(* IEC 61131-3 sources: llm-plc-st-eval/data/definitivo/qwen2.5-coder_14b/A4/few_shot, 3 files *)

(* ---- ejec_1.st ---- *)
FUNCTION_BLOCK FB_Rampa
VAR_INPUT
    SPvel : REAL; (* Consigna de velocidad *)
    paroRapido : BOOL; (* Paro rápido activo *)
    ciclo : TIME; (* Ciclo de ejecución *)
END_VAR
VAR_OUTPUT
    CVvel : REAL; (* Consigna de velocidad variable *)
END_VAR
VAR
    error : REAL; (* Error entre SPvel y CVvel *)
    dt : TIME; (* Tiempo transcurrido desde la última iteración *)
    dt_sec : REAL; (* Tiempo transcurrido en segundos *)
    rampaSubida : REAL := 10.0; (* Pendiente de subida en puntos porcentuales por segundo *)
    rampaBajada : REAL := 20.0; (* Pendiente de bajada en puntos porcentuales por segundo *)
    rampaParoRapido : REAL := 40.0; (* Pendiente de paro rápido en puntos porcentuales por segundo *)
    lastTime : TIME; (* Tiempo de la última iteración *)
END_VAR

(* Calcula el tiempo transcurrido desde la última iteración *)
dt := ciclo;
dt_sec := dt / T#1S;

(* Actualiza CVvel según las condiciones *)
IF paroRapido THEN
    (* Paro rápido activo *)
    CVvel := CVvel - rampaParoRapido * dt_sec;
    IF CVvel < 0.0 THEN
        CVvel := 0.0;
    END_IF;
ELSE
    (* Paro rápido inactivo *)
    error := SPvel - CVvel;
    IF error > 0 THEN
        (* Subida *)
        CVvel := CVvel + rampaSubida * dt_sec;
        IF CVvel > SPvel THEN
            CVvel := SPvel;
        END_IF;
    ELSE
        (* Bajada *)
        CVvel := CVvel - rampaBajada * dt_sec;
        IF CVvel < SPvel THEN
            CVvel := SPvel;
        END_IF;
    END_IF;
END_IF;

(* Actualiza el tiempo de la última iteración *)
lastTime := lastTime + ciclo;
END_FUNCTION_BLOCK

(* ---- ejec_2.st ---- *)
FUNCTION_BLOCK FB_Rampa
VAR_INPUT
    SPvel : REAL; (* Consigna de velocidad *)
    paroRapido : BOOL; (* Paro rápido activo *)
    ciclo : TIME; (* Ciclo de ejecución *)
END_VAR
VAR_OUTPUT
    CVvel : REAL; (* Condicional de velocidad *)
END_VAR
VAR
    error : REAL; (* Error entre SPvel y CVvel *)
    dt : TIME; (* Tiempo transcurrido desde la última ejecución *)
    dtSec : REAL; (* Tiempo transcurrido en segundos *)
    rampaSubida : REAL; (* Pendiente de subida *)
    rampaBajada : REAL; (* Pendiente de bajada *)
    rampaParoRapido : REAL; (* Pendiente de paro rápido *)
END_VAR

(* Inicialización de las rampas *)
rampaSubida := 10.0;
rampaBajada := 20.0;
rampaParoRapido := 40.0;

(* Cálculo del tiempo transcurrido en segundos *)
dt := ciclo;
dtSec := dt / T#1S;

(* Lógica de paro rápido *)
IF paroRapido THEN
    CVvel := MAX(0.0, CVvel - rampaParoRapido * dtSec);
ELSE
    (* Cálculo del error *)
    error := SPvel - CVvel;

    (* Ajuste de CVvel con rampa *)
    IF error > 0 THEN
        CVvel := MIN(CVvel + rampaSubida * dtSec, SPvel);
    ELSE
        CVvel := MAX(CVvel - rampaBajada * dtSec, SPvel);
    END_IF;
END_IF;

(* Evitar sobrepaso *)
IF CVvel > SPvel THEN
    CVvel := SPvel;
ELSIF CVvel < 0.0 THEN
    CVvel := 0.0;
END_IF;

END_FUNCTION_BLOCK

(* ---- ejec_3.st ---- *)
FUNCTION_BLOCK FB_Rampa
VAR_INPUT
    SPvel : REAL; (* Consigna de velocidad *)
    paroRapido : BOOL; (* Paro rápido activo *)
    ciclo : TIME; (* Ciclo de ejecución *)
END_VAR
VAR_OUTPUT
    CVvel : REAL; (* Consigna de velocidad variable *)
END_VAR
VAR
    error : REAL; (* Error entre SPvel y CVvel *)
    deltaCV : REAL; (* Cambio en CVvel *)
    rampaSubida : REAL := 10.0; (* Pendiente de subida en puntos porcentuales por segundo *)
    rampaBajada : REAL := 20.0; (* Pendiente de bajada en puntos porcentuales por segundo *)
    rampaParoRapido : REAL := 40.0; (* Pendiente de paro rápido en puntos porcentuales por segundo *)
    tiempoCiclo : TIME := T#1S; (* Tiempo de ciclo en segundos *)
END_VAR

(* Calcular el tiempo de ciclo en segundos *)
tiempoCiclo := ciclo;

(* Calcular el error *)
error := SPvel - CVvel;

(* Calcular el cambio en CVvel *)
IF paroRapido THEN
    deltaCV := rampaParoRapido * tiempoCiclo;
    IF CVvel > 0.0 THEN
        CVvel := CVvel - deltaCV;
        IF CVvel < 0.0 THEN
            CVvel := 0.0;
        END_IF
    END_IF
ELSE
    IF error > 0 THEN
        deltaCV := rampaSubida * tiempoCiclo;
    ELSE
        deltaCV := rampaBajada * tiempoCiclo;
    END_IF
    CVvel := CVvel + deltaCV;
    (* Evitar sobrepaso *)
    IF CVvel > SPvel THEN
        CVvel := SPvel;
    ELSIF CVvel < SPvel THEN
        CVvel := SPvel;
    END_IF
END_IF

END_FUNCTION_BLOCK
